(* IEC 61131-3 sources: SortJet_MasterSPS_Aufbau.fbsproj/00_Basis, 6 files *)

(* ---- StationBasisParameter.gvl ---- *)
(* METADATA
{
	"v3Meta": {
		"objectGuid": "5fda5f15-de2c-4c52-835d-2fee03387dc3"
	}
}
*)
{attribute 'allow_unqualified_access'}
NAMESPACE StationBasisParameter
// ACHTUNG: Attribute nicht ändern!
{attribute 'global_init_slot' := '310'}
VAR_GLOBAL

  starrShuttleBasisParameter                   : ARRAY [cERSTES_SHUTTLE..cLETZTES_SHUTTLE]                                OF StationBasisParameter_ST;
  starrTransfershuttleBasisParameter           : ARRAY [cERSTES_TRANSFERSHUTTLE..cLETZTES_TRANSFERSHUTTLE]                OF StationBasisParameter_ST;
  starrStationBasisParameter                   : ARRAY [cERSTE_STATION..cLETZTE_STATION]                                  OF StationBasisParameter_ST;
  starrFaecherwagenBasisParameter              : ARRAY [cERSTE_FAECHERWAGENSTATIONS_NR..cLETZTE_FAECHERWAGENSTATIONS_NR]  OF StationBasisParameter_ST;
  starrFremdanlageAuslaufStationBasisParameter : ARRAY [cERSTE_FREMDANLAGE_AUSLAUF..cLETZTE_FREMDANLAGE_AUSLAUF]          OF StationBasisParameter_ST;
  starrFremdanlageEinlaufStationBasisParameter : ARRAY [cERSTE_FREMDANLAGE_EINLAUF..cLETZTE_FREMDANLAGE_EINLAUF]          OF StationBasisParameter_ST;

END_VAR

END_NAMESPACE

(* ---- Stations_Konstanten.gvl ---- *)
(* METADATA
{
	"v3Meta": {
		"objectGuid": "55accb84-4b73-4dbf-8d20-edd3dcbc9a96"
	}
}
*)
{attribute 'allow_unqualified_access'}
NAMESPACE Stations_Konstanten
VAR_GLOBAL CONSTANT

  (* Anmerkung:
     - Konstanten die immer gleichbleiben in ihrer Benamung und nicht mehr
       angepasst werden muessen (ggf. der numerische Wert)
  *)

  // TEMPORAERE STATIONS (PLATZHALTER)
  cSTATION_DYNAMISCH       : WORD := 998;
  cSTATION_DEFAULT         : WORD := 999;
  cSTATION_TEMP            : WORD := 999;

  // Shuttle
  cSHUTTLE_101             : WORD := 101;
  cSHUTTLE_102             : WORD := 102;
  cSHUTTLE_103             : WORD := 103;
  cSHUTTLE_104             : WORD := 104;
  cSHUTTLE_105             : WORD := 105;
  cSHUTTLE_106             : WORD := 106;

  // Transfershuttle
  cSHUTTLE_150             : WORD := 150;
  cSHUTTLE_151             : WORD := 151;
  cSHUTTLE_152             : WORD := 152;
  cSHUTTLE_153             : WORD := 153;
  cSHUTTLE_154             : WORD := 154;
  cSHUTTLE_155             : WORD := 155;
  cSHUTTLE_156             : WORD := 156;
  cSHUTTLE_157             : WORD := 157;
  cSHUTTLE_158             : WORD := 158;

  // Stationen
  cSTATION_201             : WORD := 201;
  cSTATION_202             : WORD := 202;
  cSTATION_203             : WORD := 203;
  cSTATION_204             : WORD := 204;
  cSTATION_205             : WORD := 205;
  cSTATION_206             : WORD := 206;
  cSTATION_207             : WORD := 207;
  cSTATION_208             : WORD := 208;
  cSTATION_209             : WORD := 209;
  cSTATION_210             : WORD := 210;
  cSTATION_211             : WORD := 211;
  cSTATION_212             : WORD := 212;
  cSTATION_213             : WORD := 213;
  cSTATION_214             : WORD := 214;
  cSTATION_215             : WORD := 215;
  cSTATION_216             : WORD := 216;
  cSTATION_217             : WORD := 217;
  cSTATION_218             : WORD := 218;
  cSTATION_219             : WORD := 219;
  cSTATION_220             : WORD := 220;
  cSTATION_221             : WORD := 221;
  cSTATION_222             : WORD := 222;
  cSTATION_223             : WORD := 223;
  cSTATION_224             : WORD := 224;
  cSTATION_225             : WORD := 225;
  cSTATION_226             : WORD := 226;
  cSTATION_227             : WORD := 227;
  cSTATION_228             : WORD := 228;
  cSTATION_229             : WORD := 229;
  cSTATION_230             : WORD := 230;

  // Faecherwagen
  cSTATION_301             : WORD := 301;
  cSTATION_302             : WORD := 302;
  cSTATION_303             : WORD := 303;
  cSTATION_304             : WORD := 304;
  cSTATION_305             : WORD := 305;
  cSTATION_306             : WORD := 306;
  cSTATION_307             : WORD := 307;

  // Fremdanlagen
  cSTATION_401             : WORD := 401;
  cSTATION_402             : WORD := 402;
  cSTATION_403             : WORD := 403;
  cSTATION_404             : WORD := 404;

  // Einlauflinien
  cSTATION_501             : WORD := 501;
  cSTATION_502             : WORD := 502;
  cSTATION_503             : WORD := 503;

//-------------------------------------------------------------------------------------------------
// STATIONSNUMMERN [SPRECHEND]
//-------------------------------------------------------------------------------------------------
  (* Anmerkung:
     - Konstanten die immer gleichbleiben in ihrer Benamung und nicht mehr
       angepasst werden muessen (ggf. der numerische Wert)
  *)

  // Speicher
  cSPEICHER_1                 : WORD := 1;
  cSPEICHER_2                 : WORD := 2;
  cSPEICHER_3                 : WORD := 3;
  cSPEICHER_4                 : WORD := 4;
  cSPEICHER_5                 : WORD := 5;
  cSPEICHER_6                 : WORD := 6;
  cSPEICHER_7                 : WORD := 7;
  cSPEICHER_8                 : WORD := 8;

  // Fremdanlage
  cFREMDANLAGE_AUSLAUF_1      : WORD := 401;
  cFREMDANLAGE_AUSLAUF_2      : WORD := 402;
  cFREMDANLAGE_AUSLAUF_3      : WORD := 403;
  cFREMDANLAGE_AUSLAUF_4      : WORD := 404;

  cFREMDANLAGE_EINLAUF_1      : WORD := 501;
  cFREMDANLAGE_EINLAUF_2      : WORD := 502;
  cFREMDANLAGE_EINLAUF_3      : WORD := 503;

  // Hydraulik-Kreise
  cHYDRAULIKSTATION_1         : WORD := 1;
  cHYDRAULIKSTATION_2         : WORD := 2;
  cHYDRAULIKSTATION_3         : WORD := 3;

  // Wird benutzt für Horn \ Ampel
  cEINLAUFSEITE                        : WORD := 1;
  cAUSLAUFSEITE                        : WORD := 2;

  // TUEREN
  cTUER_1                              : WORD := 1;
  cTUER_2                              : WORD := 2;
  cTUER_3                              : WORD := 3;
  cTUER_4                              : WORD := 4;
  cTUER_5                              : WORD := 5;
  cTUER_6                              : WORD := 6;
  cTUER_7                              : WORD := 7;
  cTUER_8                              : WORD := 8;
  cTUER_9                              : WORD := 9;
  cTUER_10                             : WORD := 10;

  // Durchgänge Klappförderer
  cDURCHGANG_1                         : WORD := 1;
  cDURCHGANG_2                         : WORD := 2;
  cDURCHGANG_3                         : WORD := 3;

  // MMI WANDNUMMER
  //   - Wird gebraucht fuer die Fehlermeldung der Scheibenquittierung
  cMMI_WAND_1                         : WORD := 0;
  cMMI_WAND_2                         : WORD := 1;
  cMMI_WAND_3                         : WORD := 2;
  cMMI_WAND_4                         : WORD := 3;

  // HUBRAHMEN
  cHUBRAHMEN_1                        : WORD := 0;
  cHUBRAHMEN_2                        : WORD := 1;

  // ZYLINDER KENNUNG
  //   - Bei Zylinderfehlern (nicht aus-/eingefahren, Stellung ungueltig) in awFehlerInformationen[1]
  //   - Damit ist im Fehlertext erkennbar, welcher Zylinder der Station gemeint ist
  cZYLINDER_KEINE                     : WORD := 0;
  cZYLINDER_HUBRAHMEN                 : WORD := 1;
  cZYLINDER_ANSCHLAG                  : WORD := 2;
  cZYLINDER_ANSCHLAG_HORIZONTAL       : WORD := 3;
  cZYLINDER_ABSCHRANKUNG              : WORD := 4;
  cZYLINDER_DICKENVERSTELLUNG         : WORD := 5;
  cZYLINDER_ROELLCHENLEISTE           : WORD := 6;
  cZYLINDER_WANDVERSTELLUNG           : WORD := 7;
  cZYLINDER_QUERACHSE                 : WORD := 8;
  cZYLINDER_ARRETIERUNG               : WORD := 9;
  cZYLINDER_GREIFER_HUB               : WORD := 10;
  cZYLINDER_ZANGE_EINLAUF             : WORD := 11;
  cZYLINDER_ZANGE_AUSLAUF             : WORD := 12;

  // EBENEN
  cEBENE_1                            : WORD := 2#0000000000000001; // 1;
  cEBENE_2                            : WORD := 2#0000000000000010; // 2;

END_VAR

END_NAMESPACE

(* ---- Initialisierung.prg.st ---- *)
(* METADATA
{
	"v3Meta": {
		"objectGuid": "cf26b0b7-1f73-4db7-a5c7-b5425b79f88d"
	}
}
*)
PROGRAM Initialisierung
VAR_INPUT

  // BOOL
  bpReset                             : BOOL;
  bpInitialisierung                   : BOOL;

END_VAR
VAR_OUTPUT

  // BOOL
  bpFehler                             : BOOL;
  bpInitialisierungAktiv               : BOOL;

END_VAR
VAR

  // BOOL
  blErsterZyklus                       : BOOL := TRUE;
  blReturn                             : BOOL; // Wird gesetzt um im nächsten Zyklus mit Return rauszuspringen. Vorher sollen die WatchIO's zurück gesetzt werden
  blFreigabeZumReferenzieren           : BOOL;
  blFreigabeAutokreis                  : BOOL;
  blAlleSKGeschlossen                  : BOOL;
  blDruckluftOK                        : BOOL;
  blShuttleErreichbar                  : BOOL;
  blInitDurchFehlerGeblockt            : BOOL;

  // WORD
  wlIndex                              : WORD;
  wlSubIndex                           : WORD;
  wlMeldungsnummer                     : WORD;

  // INT
  ilAnzahlStationenReferenzAktiv       : INT;
  ilAnzahlShuttleReferenzAktiv         : INT;
  ilAnzahlTransfershuttleReferenzAktiv : INT;

  // TIMER
  tonlWait_Init                        : TON;
  tonlFreigabeReferenzierung           : TON;

  // STEPS
  steplInitialisierung                 : STEPS_TE;

END_VAR

//-------------------------------------------------------------------------------------------------
// INITIALISIERUNG
//-------------------------------------------------------------------------------------------------
IF ( blErsterZyklus ) THEN
  blErsterZyklus := FALSE;
END_IF

IF bgInitialisierungUeberbruecken THEN
  M_Init_Ok := TRUE;
END_IF

IF (  NOT M_Init_Ok
     AND NOT blErsterZyklus )
THEN
  bpInitialisierung := TRUE;
  blReturn          := FALSE;
ELSIF blReturn THEN
  RETURN; // Init abgeschlossen
ELSE
  bpInitialisierung := FALSE;
  blReturn          := TRUE;
END_IF

//-------------------------------------------------------------------------------------------------
// AKTIONEN
//-------------------------------------------------------------------------------------------------
Meldungen();
Init();

//-------------------------------------------------------------------------------------------------
// Setzen der Freigabe für die Initialisierung ( Referenzierung )
//-------------------------------------------------------------------------------------------------
// Abfrage ob kein Reset aktiv ist
blFreigabeAutokreis := TRUE;
FOR wlIndex := cERSTER_AUTOMATIKKREIS TO cLETZTER_AUTOMATIKKREIS DO
  IF agbResetAktiv[wlIndex] THEN
    blFreigabeAutokreis := FALSE;
  END_IF
END_FOR

blInitDurchFehlerGeblockt := FALSE;
FOR wlIndex := cERSTER_AUTOMATIKKREIS TO cLETZTER_AUTOMATIKKREIS DO
  blInitDurchFehlerGeblockt := blInitDurchFehlerGeblockt OR Job.ablFehlerAktiv[wlIndex];
END_FOR

blFreigabeZumReferenzieren := ( (     NotHalt.bpNotHaltOK
                                  AND blAlleSKGeschlossen )
                                OR bgSicherheitstechnikBruecken )
                              AND ( bgMMIOK OR bgMMIBruecken )
                              AND blDruckluftOK
                              AND blShuttleErreichbar
                              AND blFreigabeAutokreis
                              AND bgEtherCatOK
                              AND NOT blInitDurchFehlerGeblockt;

tonlFreigabeReferenzierung(IN := blFreigabeZumReferenzieren ,PT := t#5s);
END_PROGRAM

(* ---- Main.prg.st ---- *)
(* METADATA
{
	"v3Meta": {
		"objectGuid": "38b1ebdf-93dc-4d21-adff-5cd8952a9cb8"
	}
}
*)
PROGRAM Main
VAR

  // BOOL
  blErsterZyklus : BOOL := TRUE;
  blZweiterZyklus : BOOL := FALSE;

  aStation1Wand : ARRAY[cWAND_1..cANZAHL_WAENDE] OF BOOL;
  aStation2Wand : ARRAY[cWAND_1..cANZAHL_WAENDE] OF BOOL;

  // BLINK
  Flasher02                  : BLINK;
  Flasher03                  : BLINK;
  Flasher05                  : BLINK;
  Flasher10                  : BLINK;
  Flasher12                  : BLINK;

  // WORD
  wlIndex                    : WORD;

  // TRIGGER
  rtlChangeWatchIOStatus     : R_TRIG;

  // Events
  sCallbackOnlineChange      : CB.CB_CALLBACK;
  peCallbackStopOnlineChange : CB.ERROR;

END_VAR

VAR_OUTPUT

  // TRIGGER
  rtlEtherCatOK              : R_TRIG;
END_VAR
// -------------------------------------------------------------------------
// -----!!! Vor dem Befehl <MsgBegin> sollte keine Anweisung stehen !!!-----
TCPMain.l_fb_SortjetHMI.MsgBegin();
// -----!!! Vor dem Befehl <MsgBegin> sollte keine Anweisung stehen !!!-----
// -------------------------------------------------------------------------

TCPMain();

EtherCAT_Master.StartConfigWithLessDevice := TRUE;

IF ( Auftraege.bgInbetriebnahmeAblaeufe ) THEN
  Auftraege();
END_IF

Flasher();
Merker();

//EventsRegistrieren();
CheckReset();
StationBasisZuweisungen();
Auftraege();
Interface_SLC();
NotHalt();
SteuerungSicherheitskreise();
Stop_Baustein();
Initialisierung();
SystemCheck();
Job();
StationsAufrufe();

IF ( blZweiterZyklus ) THEN
  blZweiterZyklus := FALSE;
  StartUpCheck();
END_IF

IF ( blErsterZyklus ) THEN
  blErsterZyklus := FALSE;
  blZweiterZyklus := TRUE;
  // !!! Muss NACH dem Aufruf von Job erfolgen, da sonst die MKs nicht initialisiert sind !!!
  wgAnzahlSystemcheckZyklen := getAnzahlSystemcheckZyklen();
END_IF

StatusAnlage();
Visu();

(* Hinweis:
   - Schrittketten Auswertung
*)
Schrittketten_Logger();
AntriebeVerfahren();

bgMMIOK := TCPMain.l_fb_SortjetHMI.o_b_WatchdogOk;
// -------------------------------------------------------------------------
// -!!! Nach dem Befehl <MsgEnd> sollte keine weitere Anweisung folgen !!!--
TCPMain.l_fb_SortjetHMI.MsgEnd();
// -!!! Nach dem Befehl <MsgEnd> sollte keine weitere Anweisung folgen !!!--
// -------------------------------------------------------------------------
END_PROGRAM

(* ---- SlowTask.prg.st ---- *)
(* METADATA
{
	"v3Meta": {
		"objectGuid": "14e1f1f9-a11c-4000-82c5-ba9f94dc3c1b"
	}
}
*)
PROGRAM SlowTask
VAR

  // EtherCAT Reset
  bpSlave                    : POINTER TO ETCSlave;

  // BOOL
  blECatOK                   : BOOL;
  blRestartEtherCatMMI       : BOOL;

  // STEPS
  steplEtherCat_Restart      : Steps_TE;

  // TIMER
  tonlWaitInit               : TON;
  tonl_Step                  : TON;
  tonlEtherCat_Start_TimeOut : TON;

  // TRIGGER
  rtrigECatOK                : R_TRIG;
END_VAR

StationBasisZuweisungen.M_AufrufeZuweisungen();
EtherCAT_Restart();
END_PROGRAM

(* ---- StatusAnlage.prg.st ---- *)
(* METADATA
{
	"v3Meta": {
		"objectGuid": "008eb84c-ed0d-4cb0-9376-462b0a38bc1c"
	}
}
*)
PROGRAM StatusAnlage
VAR

  // WORD
  wlIndex          : WORD;

END_VAR
VAR_OUTPUT

  // BOOLEAN
  abpDruckluftOK    : ARRAY [cERSTER_AUTOMATIKKREIS..cLETZTER_AUTOMATIKKREIS] OF BOOL;
  bpAnlageOK        : BOOL;
END_VAR
VAR

  // TIMER
  toflDruckluftShuttleOK           : ARRAY[cERSTES_SHUTTLE..cLETZTES_SHUTTLE] OF TOF;
  toflDruckluftTSShuttleOK         : ARRAY[cERSTES_TRANSFERSHUTTLE..cLETZTES_TRANSFERSHUTTLE] OF TOF;
  toflDruckluft101_OK              : TOF;
  toflDruckluft102_OK              : TOF;
  toflDruckluftFW_OK               : TOF;
  toflDruckluftAnlegetisch201_OK   : TOF;
  toflDruckluftAnlegetisch205_OK   : TOF;

END_VAR

VAR

  // Druckluft
  in_bDruckluft_FW_OK                                  : BOOL; // Wartungseinheit
  in_bDruckluft_101_OK                        AT %I*   : BOOL; // Wartungseinheit
  in_bDruckluft_102_OK                        AT %I*   : BOOL; // Wartungseinheit

  // CAB 2
  in_bCAB2_KlimaGeraet_OK                     AT %I* : BOOL;
  in_bCAB2_LS_Netzteil_24V_OK                 AT %I* : BOOL;
  in_bCAB2_LS_24V_Schaltschrank_OK            AT %I* : BOOL;
  in_bCAB2_LS_24V_Boxen_OK                    AT %I* : BOOL;
  in_bCAB2_LS_400V_OK                         AT %I* : BOOL;
  in_bCAB2_LS_Netzfilter_400V_OK              AT %I* : BOOL;
  in_bCAB2_LS_230V_OK                         AT %I* : BOOL;
  in_bCAB2_Sicherheitsrelais_201_Kippen_OK    AT %I* : BOOL; // Sicherheitsrelais 201 Hydraulik / kippen OK

END_VAR

VAR CONSTANT

  // TIME
  ZEIT_DRUCKWAECHTERSIGNAL_ENTPRELLT : TIME := T#3s;

END_VAR
//-------------------------------------------------------------------------------------------------
// STATUS DER BASIS-KOMPONENTEN INHERHALB DER ANLAGE
//-------------------------------------------------------------------------------------------------

// Entprellen des Druckwaechter- Einheit => SHUTTLE
FOR wlIndex := cERSTES_SHUTTLE TO cLETZTES_SHUTTLE DO
  toflDruckluftShuttleOK[wlIndex]( IN := aShuttle[wlIndex].in_bDruckluft_OK OR starrShuttleBasisParameter[wlIndex].stMKs.bDeaktivieren ,
                                   PT := ZEIT_DRUCKWAECHTERSIGNAL_ENTPRELLT );
END_FOR

// Entprellen des Druckwaechter- Einheit => TRANSFERSHUTTLE
FOR wlIndex := cERSTES_TRANSFERSHUTTLE TO cLETZTES_TRANSFERSHUTTLE DO
  toflDruckluftTSShuttleOK[wlIndex]( IN := aTransfershuttles[wlIndex].in_bDruckluftWartungseinheitOK OR starrTransfershuttleBasisParameter[wlIndex].stMKs.bDeaktivieren ,
                                     PT := ZEIT_DRUCKWAECHTERSIGNAL_ENTPRELLT );
END_FOR

// Entprellen des Druckwaechters => ANLEGETISCH
toflDruckluftAnlegetisch201_OK( IN := Globale_Bausteine.Anlegetisch201.in_bDruckluft_OK OR starrStationBasisParameter[cSTATION_201].stMKs.bDeaktivieren OR NOT starrStationBasisParameter[cSTATION_201].stMKs.stStationsAufbau.bDruckluft ,
                                PT := ZEIT_DRUCKWAECHTERSIGNAL_ENTPRELLT );
toflDruckluftAnlegetisch205_OK( IN := Globale_Bausteine.Anlegetisch205.in_bDruckluft_OK OR starrStationBasisParameter[cSTATION_205].stMKs.bDeaktivieren OR NOT starrStationBasisParameter[cSTATION_205].stMKs.stStationsAufbau.bDruckluft ,
                                PT := ZEIT_DRUCKWAECHTERSIGNAL_ENTPRELLT );

toflDruckluft101_OK( In := in_bDruckluft_101_OK, PT := ZEIT_DRUCKWAECHTERSIGNAL_ENTPRELLT );
toflDruckluft102_OK( In := in_bDruckluft_102_OK, PT := ZEIT_DRUCKWAECHTERSIGNAL_ENTPRELLT );
toflDruckluftFW_OK( In := in_bDruckluft_FW_OK OR %MX1.1, PT := ZEIT_DRUCKWAECHTERSIGNAL_ENTPRELLT ); // TODO wenn Wartungseinheit verbaut

// Auswertung und hier pruefen ob Betriebsstopp ausgeloest werden muss
// AK1 = Foerderstrecke (201 - 208), Shuttle 101 und die Transfershuttles (151, 152)
abpDruckluftOK[cAUTOMATIKKREIS_1] := (   ( toflDruckluftShuttleOK[cSHUTTLE_101].Q OR starrShuttleBasisParameter[cSHUTTLE_101].stMKs.bDeaktivieren OR NOT starrShuttleBasisParameter[cSHUTTLE_101].stMKs.stStationsAufbau.bDruckluft )
                                       AND toflDruckluft101_OK.Q
                                       AND toflDruckluftAnlegetisch201_OK.Q
                                       AND toflDruckluftAnlegetisch205_OK.Q
                                       AND ( toflDruckluftTSShuttleOK[cSHUTTLE_151].Q OR starrTransfershuttleBasisParameter[cSHUTTLE_151].stMKs.bDeaktivieren)
                                       AND ( toflDruckluftTSShuttleOK[cSHUTTLE_152].Q OR starrTransfershuttleBasisParameter[cSHUTTLE_152].stMKs.bDeaktivieren)
                                     ) OR bgInbetriebnahmeBit;

// AK2 = Shuttle 102, Transfershuttles (151, 152) und Faecherwagen (301 - 305)
abpDruckluftOK[cAUTOMATIKKREIS_2] := (   ( toflDruckluftShuttleOK[cSHUTTLE_102].Q OR starrShuttleBasisParameter[cSHUTTLE_102].stMKs.bDeaktivieren OR NOT starrShuttleBasisParameter[cSHUTTLE_102].stMKs.stStationsAufbau.bDruckluft )
                                       AND toflDruckluft102_OK.Q
                                       AND toflDruckluftFW_OK.Q
                                       AND ( toflDruckluftTSShuttleOK[cSHUTTLE_151].Q OR starrTransfershuttleBasisParameter[cSHUTTLE_151].stMKs.bDeaktivieren)
                                       AND ( toflDruckluftTSShuttleOK[cSHUTTLE_152].Q OR starrTransfershuttleBasisParameter[cSHUTTLE_152].stMKs.bDeaktivieren)
                                     ) OR bgInbetriebnahmeBit;

bpAnlageOK := ( ( in_bCAB2_LS_Netzteil_24V_OK
                  AND in_bCAB2_LS_24V_Schaltschrank_OK
                  AND in_bCAB2_LS_24V_Boxen_OK
                  AND in_bCAB2_LS_400V_OK
                  AND in_bCAB2_LS_Netzfilter_400V_OK )
                OR bgInbetriebnahmeBit) ;

// Meldungen CAB 2
WatchIo(NOT bgInbetriebnahmeBit AND NOT in_bCAB2_KlimaGeraet_OK,  ioccCAB2_Klimageraet_Nicht_OK);
WatchIo(NOT in_bCAB2_LS_Netzteil_24V_OK,                          ioccCAB2_Netzteil_24V_Nicht_Ok);
WatchIo(NOT in_bCAB2_LS_24V_Schaltschrank_OK,                     ioccCAB2_LS_24V_Schaltschrank_Nicht_OK);
WatchIo(NOT in_bCAB2_LS_24V_Boxen_OK,                             ioccCAB2_LS_24V_Boxen_Nicht_OK);
WatchIo(NOT in_bCAB2_LS_400V_OK,                                  ioccCAB2_LS_400V_Nicht_OK_);
WatchIo(NOT in_bCAB2_LS_Netzfilter_400V_OK,                       ioccCAB2_LS_Netzfilter_400V_Nicht_OK);
WatchIo(NOT in_bCAB2_Sicherheitsrelais_201_Kippen_OK,             ioccCAB2_Sicherheitsrelais_201_Kippen_Nicht_OK);
WatchIo(NOT in_bCAB2_LS_230V_OK,                                  ioccCAB2_LS_230V_Nicht_OK);

WatchIo(NOT bgInbetriebnahmeBit AND NOT toflDruckluft101_OK.Q,  ioccDruckluft1);
WatchIo(NOT bgInbetriebnahmeBit AND NOT toflDruckluft102_OK.Q,  ioccDruckluft2);
WatchIo(NOT bgInbetriebnahmeBit AND NOT toflDruckluftFW_OK.Q,   ioccDruckluft3);
END_PROGRAM
